Fanuc KAREL source: kb00019.KL

-- PROVISIONAL review KL for V770-1; original PC SHA256 cf23be6e8903fe6563f7ef4f0a2544f0dc706da0e7402aceb4a09f75d0cdefa0
-- Incomplete behavior may be omitted. Consult companion uncertainty JSON. Do not deploy.
PROGRAM KB00019
%NOLOCKGROUP
BEGIN
  -- UNRESOLVED_PC offsets 5-14; opcodes 3F,75
  -- UNRESOLVED_PC offsets 19-26; opcodes 9D,23
  -- UNRESOLVED_PC offsets 31-49; opcodes 27,22,2A,22,31
  -- UNRESOLVED_PC offsets 54-58; opcodes 7F
END KB00019
